(* IEC 61131-3 sources: kns-pump-station/tests/POUs/Station/FB_PowerRestore_Test, 14 files *)

(* ---- DemandRisingAfterDelayKeepsSequence.method.decl.st ---- *)
// 04 §13.2, PMI-34: после задержки потребность растёт (ступенчатый автомат после Restart начинает с нуля и
// подтверждает второй насос позже конца задержки) — последовательность не завершается, пока не пущены все
// запрошенные: подпорный — через tSeqStep после подтверждения ведущего, событие 101010 со значением 2
METHOD PRIVATE DemandRisingAfterDelayKeepsSequence
VAR
    fbDut  : FB_PowerRestore;           // ФБ под тестом
    fbTime : PL.FB_FakeTime;            // подменное время, старт 1 ч
    stCfg  : ST_StationCfg;             // уставки по умолчанию: tPlcStart 10 с, tPwrRestart 10 с, tSeqStep 15 с
    fbSink : FB_FakeEventSink;          // подменный журнал
END_VAR

(* ---- FirstCallIgnoresPowerInput.method.decl.st ---- *)
// DESIGN 6.9: в первом вызове вход ES301 ещё не посчитан устройством — пропадание не фиксируется; со второго
// вызова — да
METHOD PRIVATE FirstCallIgnoresPowerInput
VAR
    fbDut  : FB_PowerRestore;           // ФБ под тестом
    fbTime : PL.FB_FakeTime;            // подменное время, старт 1 ч
    stCfg  : ST_StationCfg;             // уставки по умолчанию: tPlcStart 10 с, tPwrRestart 10 с, tSeqStep 15 с
    fbSink : FB_FakeEventSink;          // подменный журнал
END_VAR

(* ---- LastStepUnconfirmedFinishesOnTimeout.method.decl.st ---- *)
// 04 §13.2: пуск последнего нужного шага не подтвердился (насос отказал, замены нет) — последовательность
// завершается через STN_SEQ_START_TIMEOUT, а не держит Restart бесконечно
METHOD PRIVATE LastStepUnconfirmedFinishesOnTimeout
VAR
    fbDut  : FB_PowerRestore;           // ФБ под тестом
    fbTime : PL.FB_FakeTime;            // подменное время, старт 1 ч
    stCfg  : ST_StationCfg;             // уставки по умолчанию: tPlcStart 10 с, tPwrRestart 10 с, tSeqStep 15 с
    fbSink : FB_FakeEventSink;          // подменный журнал
END_VAR

(* ---- NothingRequiredFinishesImmediately.method.decl.st ---- *)
// 04 §13.2: насосы не нужны — последовательность завершается сразу после задержки (101010 со значением 0)
METHOD PRIVATE NothingRequiredFinishesImmediately
VAR
    fbDut  : FB_PowerRestore;           // ФБ под тестом
    fbTime : PL.FB_FakeTime;            // подменное время, старт 1 ч
    stCfg  : ST_StationCfg;             // уставки по умолчанию: tPlcStart 10 с, tPwrRestart 10 с, tSeqStep 15 с
    fbSink : FB_FakeEventSink;          // подменный журнал
END_VAR

(* ---- PlcStartDelaysAllRequests.method.decl.st ---- *)
// 04 §13.3, PMI-01, PMI-35: старт ПЛК — «задержка» tPlcStart = 10 с без запросов (событие 101009), затем первый
// шаг
METHOD PRIVATE PlcStartDelaysAllRequests
VAR
    fbDut  : FB_PowerRestore;           // ФБ под тестом
    fbTime : PL.FB_FakeTime;            // подменное время, старт 1 ч
    stCfg  : ST_StationCfg;             // уставки по умолчанию: tPlcStart 10 с, tPwrRestart 10 с, tSeqStep 15 с
    fbSink : FB_FakeEventSink;          // подменный журнал
END_VAR

(* ---- PowerLossBlocksRequests.method.decl.st ---- *)
// 04 §13.1, PMI-33: нет напряжения — PowerLost, запросов нет, событие 101008
METHOD PRIVATE PowerLossBlocksRequests
VAR
    fbDut  : FB_PowerRestore;           // ФБ под тестом
    fbTime : PL.FB_FakeTime;            // подменное время, старт 1 ч
    stCfg  : ST_StationCfg;             // уставки по умолчанию: tPlcStart 10 с, tPwrRestart 10 с, tSeqStep 15 с
    fbSink : FB_FakeEventSink;          // подменный журнал
END_VAR

(* ---- PowerLossDuringSequenceRestarts.method.decl.st ---- *)
// 04 §13.2: пропадание напряжения во время последовательного пуска — с начала: задержка и первый шаг
METHOD PRIVATE PowerLossDuringSequenceRestarts
VAR
    fbDut  : FB_PowerRestore;           // ФБ под тестом
    fbTime : PL.FB_FakeTime;            // подменное время, старт 1 ч
    stCfg  : ST_StationCfg;             // уставки по умолчанию: tPlcStart 10 с, tPwrRestart 10 с, tSeqStep 15 с
    fbSink : FB_FakeEventSink;          // подменный журнал
END_VAR

(* ---- RestoreWaitsTPwrRestart.method.decl.st ---- *)
// 04 §13.2, PMI-34: напряжение вернулось — «задержка» tPwrRestart = 10 с (событие 101009), затем первый шаг
METHOD PRIVATE RestoreWaitsTPwrRestart
VAR
    fbDut  : FB_PowerRestore;           // ФБ под тестом
    fbTime : PL.FB_FakeTime;            // подменное время, старт 1 ч
    stCfg  : ST_StationCfg;             // уставки по умолчанию: tPlcStart 10 с, tPwrRestart 10 с, tSeqStep 15 с
    fbSink : FB_FakeEventSink;          // подменный журнал
END_VAR

(* ---- Run.method.decl.st ---- *)
// Помощник: uiSteps шагов времени tStep; входы ФБ тест задаёт присваиванием
METHOD PRIVATE Run
VAR_IN_OUT
    fbDut  : FB_PowerRestore;           // ФБ под тестом
    fbTime : PL.FB_FakeTime;            // подменное время
    stCfg  : ST_StationCfg;             // уставки
END_VAR
VAR_INPUT
    tStep   : TIME;                     // шаг времени
    uiSteps : UINT;                     // шагов
END_VAR
VAR
    uiStep : UINT;                      // номер шага
END_VAR

(* ---- Run.method.impl.st ---- *)
FOR uiStep := 1 TO uiSteps DO
    fbTime.Advance(tStep := tStep);
    fbDut(itfTime := fbTime, stCfg := stCfg);
END_FOR

(* ---- SeqRemainCountsDown.method.decl.st ---- *)
// 04 §13.2, PMI-34: uiSeqRemain_s — остаток до следующего шага в целых секундах вверх
METHOD PRIVATE SeqRemainCountsDown
VAR
    fbDut  : FB_PowerRestore;           // ФБ под тестом
    fbTime : PL.FB_FakeTime;            // подменное время, старт 1 ч
    stCfg  : ST_StationCfg;             // уставки по умолчанию: tPlcStart 10 с, tPwrRestart 10 с, tSeqStep 15 с
    fbSink : FB_FakeEventSink;          // подменный журнал
END_VAR

(* ---- SequenceOnePumpPerStep.method.decl.st ---- *)
// 04 §13.2, PMI-34: шаги по одному насосу — следующий через tSeqStep = 15 с после подтверждения пуска; конец — все
// запрошенные пущены, событие 101010 с числом пущенных
METHOD PRIVATE SequenceOnePumpPerStep
VAR
    fbDut  : FB_PowerRestore;           // ФБ под тестом
    fbTime : PL.FB_FakeTime;            // подменное время, старт 1 ч
    stCfg  : ST_StationCfg;             // уставки по умолчанию: tPlcStart 10 с, tPwrRestart 10 с, tSeqStep 15 с
    fbSink : FB_FakeEventSink;          // подменный журнал
END_VAR

(* ---- StepAdvancesOnTimeoutIfStartFails.method.decl.st ---- *)
// 04 §13.2: пуск шага не подтвердился (АВР назначил замену) — следующий шаг через STN_SEQ_START_TIMEOUT = 30 с
METHOD PRIVATE StepAdvancesOnTimeoutIfStartFails
VAR
    fbDut  : FB_PowerRestore;           // ФБ под тестом
    fbTime : PL.FB_FakeTime;            // подменное время, старт 1 ч
    stCfg  : ST_StationCfg;             // уставки по умолчанию: tPlcStart 10 с, tPwrRestart 10 с, tSeqStep 15 с
    fbSink : FB_FakeEventSink;          // подменный журнал
END_VAR

(* ---- TimeBackwardsRestartsDelay.method.decl.st ---- *)
// Время назад — задержка tPlcStart начинается заново, раннего пуска нет
METHOD PRIVATE TimeBackwardsRestartsDelay
VAR
    fbDut  : FB_PowerRestore;           // ФБ под тестом
    fbTime : PL.FB_FakeTime;            // подменное время, старт 1 ч
    stCfg  : ST_StationCfg;             // уставки по умолчанию: tPlcStart 10 с, tPwrRestart 10 с, tSeqStep 15 с
    fbSink : FB_FakeEventSink;          // подменный журнал
END_VAR
